(*
SPDX-FileCopyrightText: © 2026 Oleksandr Tiutyk <trofimich@gmail.com>
SPDX-License-Identifier: MIT
License: https://opensource.org/license/mit
*)

(*!
<summary>
Beckhoff EL5151: 1-channel incremental encoder interface terminal (24 V HTL, single-ended).
</summary>
<description>
Represents Standard 32-bit (MDP 511) main PDOs: TxPDO 0x1A00 and RxPDO 0x1600.
Ch1 contains 16-bit status/control and 32-bit counter, latch and preset values.
Optional period/frequency/timestamp PDOs are outside this model; disable or link them separately.
The Standard 16-bit process image is unsupported.
When used for I/O, link located fields or their containing buffers to the matching selected PDOs.
The record is not a packed wire buffer; compiler padding is not part of the device specification.
Unlinked/default values do not prove valid I/O. The caller evaluates bus/channel validity before use.
Use one owner task per instance and externally synchronize other access; multi-field snapshots are not atomic.
Copies store data without creating hardware links. Keep borrowed field references valid while consumers are bound.
This passive record performs no validation, synchronization, configuration or protocol advancement.
</description>
*)
TYPE EL5151 :
STRUCT
	Ch1 : INCREMENTAL_ENCODER_CHANNEL;
END_STRUCT
END_TYPE

(* stored: Version 1.1.0.1, ProductVersion 3.1.4026.20
   DUT EL5151: Id {201ad3a3-6b20-4989-b6bd-74d7b5b281ad} *)
